(* IEC 61131-3 sources: Test-Git_ESME26/TestProgettoESME_26.fbsproj/PacDriveLib Migration/Motion/MultiCam/PDL_FB_MultiCam.fb.st^/PlcOpen, 3 files *)

(* ---- CallPLCopenFBs.meth.st ---- *)
METHOD PRIVATE CallPLCopenFBs : BOOL
VAR_INPUT
END_VAR

(*********************************************************************************************************************)
fbMoveAbsolute();

IF fbMoveAbsolute.Error THEN
	SetDiagOutput(	i_etDiag	:= GD.ET_Diag.UnexpectedProgramBehavior,
					i_etDiagExt := PDL_ET_DiagExt.UnexpectedFeedback,
					i_sMsg		:= CONCAT('MC_MoveAbsolute.ErrorID: ', PLCO.FC_EtResultToString(fbMoveAbsolute.ErrorID) ));
	fbMoveAbsolute.Execute := FALSE;

	q_xReady		:= FALSE;
	q_xSynActive	:= FALSE;
	q_xXLowEnd		:= FALSE;
	q_xXHighEnd		:= FALSE;
	q_xInWSWindow	:= FALSE;
	etState := ET_MulticamState.controllerStop;
END_IF

(*********************************************************************************************************************)
fbCamIn();

IF fbCamIn.Error THEN

	SetDiagOutput(	i_etDiag	:= GD.ET_Diag.UnexpectedProgramBehavior,
					i_etDiagExt := PDL_ET_DiagExt.UnexpectedFeedback,
					i_sMsg		:= CONCAT('MC_CamIn.ErrorID: ', PLCO.FC_EtResultToString(fbCamIn.ErrorID) ));

	fbCamIn.Execute := FALSE;
	q_xReady		:= FALSE;
	q_xSynActive	:= FALSE;
	q_xXLowEnd		:= FALSE;
	q_xXHighEnd		:= FALSE;
	q_xInWSWindow	:= FALSE;
	etState := ET_MulticamState.controllerStop;
END_IF

(*********************************************************************************************************************)
fbCamIn2();

IF fbCamIn2.Error THEN

	SetDiagOutput(	i_etDiag	:= GD.ET_Diag.UnexpectedProgramBehavior,
					i_etDiagExt := PDL_ET_DiagExt.UnexpectedFeedback,
					i_sMsg		:= CONCAT('MC_CamIn.ErrorID: ', PLCO.FC_EtResultToString(fbCamIn2.ErrorID) ));

	fbCamIn2.Execute := FALSE;
	q_xReady		:= FALSE;
	q_xSynActive	:= FALSE;
	q_xXLowEnd		:= FALSE;
	q_xXHighEnd		:= FALSE;
	q_xInWSWindow	:= FALSE;
	etState := ET_MulticamState.controllerStop;
END_IF

(*********************************************************************************************************************)

xCamInInSync :=    fbCamIn.InSync
			   AND NOT xCamIn2Active
			   OR  fbCamIn2.InSync
			   AND xCamIn2Active;

xCamInEndOfProfile :=      fbCamIn.EndOfProfile
					   AND NOT xCamIn2Active
					   OR  fbCamIn2.EndOfProfile
					   AND xCamIn2Active;

(* ---- SetPosition.meth.st ---- *)
METHOD PRIVATE SetPosition : BOOL
VAR_INPUT
	i_ifAxis		: MOIN.IF_Axis;
	i_lrPosition	: LREAL;
	i_xRelative		: BOOL;
END_VAR

VAR
	etSetPosResult				: PLCO.ET_Result;
END_VAR

SetPosition := TRUE;

fbSetPos( Execute		:= FALSE );
fbSetPos(	Axis		:= i_ifAxis,
			Execute		:= TRUE,
			Position	:= i_lrPosition,
			Relative	:= i_xRelative,
			ErrorId		=> etSetPosResult );

IF etSetPosResult <> PLCO.ET_Result.Ok THEN

	SetDiagOutput(	i_etDiag	:= GD.ET_Diag.UnexpectedProgramBehavior,
					i_etDiagExt := PDL_ET_DiagExt.UnexpectedFeedback,
					i_sMsg		:= CONCAT('MC_SetPosition: ', TO_STRING(etSetPosResult)));

	SetPosition := FALSE;//no success

	etState := ET_MulticamState.controllerStop;
END_IF

(* ---- StartCam.meth.st ---- *)
METHOD PRIVATE StartCam : BOOL
VAR_INPUT
	i_etBufferMode 			: PLCO.MC_Buffer_Mode;
	i_stMultiCamData		: PDL_ST_MultiCam;
	i_lrMasterStartPosition	: LREAL := 0;
	i_xPeriodic 			: BOOL := TRUE;
	i_etMasterStartMode		: PLCO.MC_Master_Start_Mode := PLCO.MC_Master_Start_Mode.Absolute;
	i_etSlaveStartMode		: PLCO.MC_Slave_Start_Mode := PLCO.MC_Slave_Start_Mode.RampIn;
	i_xInputVelocity		: BOOL := FALSE;
	i_etDirection			: PLCO.MC_Direction := PLCO.MC_Direction.ShortestWay;
END_VAR

IF xCamIn2Active THEN

	//camIn1
	//***********************************************************************************
	xCamIn2Active := FALSE;
	fbCamIn2( Execute := FALSE );

	IF i_xInputVelocity THEN
		fbCamIn.VelocityOffsetRampIn		:= i_lrWSVel;
		fbCamIn.AccelerationOffsetRampIn	:= i_lrWSAcc;
		fbCamIn.DecelerationOffsetRampIn	:= i_lrWSAcc;
		fbCamIn.JerkOffsetRampIn			:= i_lrWsJerk;
	ELSE
		IF ifDriveConfig <> 0 THEN
			IF ifDriveConfig.MaxVel <> 0 THEN
				fbCamIn.VelocityOffsetRampIn		:= ifDriveConfig.MaxVel;
			ELSE
				fbCamIn.VelocityOffsetRampIn		:= lrLimitMaxVel;
			END_IF

			IF ifDriveConfig.MaxAcc <> 0 THEN
				fbCamIn.AccelerationOffsetRampIn	:= ifDriveConfig.MaxAcc;
				fbCamIn.DecelerationOffsetRampIn	:= ifDriveConfig.MaxAcc;
			ELSE
				fbCamIn.AccelerationOffsetRampIn	:= lrLimitMaxAccDec;
				fbCamIn.DecelerationOffsetRampIn	:= lrLimitMaxAccDec;
			END_IF
		ELSE
			fbCamIn.VelocityOffsetRampIn		:= lrLimitMaxVel;
			fbCamIn.AccelerationOffsetRampIn	:= lrLimitMaxAccDec;
			fbCamIn.DecelerationOffsetRampIn	:= lrLimitMaxAccDec;
		END_IF
		fbCamIn.JerkOffsetRampIn			:= 0;
	END_IF

	fbCamIn(	Execute						:= TRUE,
				CamTableID					:= i_stMultiCamData,
				BufferMode					:= i_etBufferMode,
				Periodic					:= i_xPeriodic,
				MasterOffset				:= 0,
				SlaveOffset					:= 0,
				MasterScaling				:= 1,
				SlaveScaling				:= 1,
				MasterStartMode				:= i_etMasterStartMode,
				SlaveStartMode				:= i_etSlaveStartMode,
				RampInDirection				:= i_etDirection,
				MasterStartPosition			:= i_lrMasterStartPosition);

ELSE
	//camIn2
	//***********************************************************************************
	xCamIn2Active := TRUE;
	fbCamIn( Execute := FALSE );

	IF i_xInputVelocity THEN
		fbCamIn2.VelocityOffsetRampIn		:= i_lrWSVel;
		fbCamIn2.AccelerationOffsetRampIn	:= i_lrWSAcc;
		fbCamIn2.DecelerationOffsetRampIn	:= i_lrWSAcc;
		fbCamIn2.JerkOffsetRampIn			:= i_lrWsJerk;
	ELSE
		IF ifDriveConfig <> 0 THEN
			IF ifDriveConfig.MaxVel <> 0 THEN
				fbCamIn2.VelocityOffsetRampIn		:= ifDriveConfig.MaxVel;
			ELSE
				fbCamIn2.VelocityOffsetRampIn		:= lrLimitMaxVel;
			END_IF
			IF ifDriveConfig.MaxAcc <> 0 THEN
				fbCamIn2.AccelerationOffsetRampIn	:= ifDriveConfig.MaxAcc;
				fbCamIn2.DecelerationOffsetRampIn	:= ifDriveConfig.MaxAcc;
			ELSE
				fbCamIn2.AccelerationOffsetRampIn	:= lrLimitMaxAccDec;
				fbCamIn2.DecelerationOffsetRampIn	:= lrLimitMaxAccDec;
			END_IF
		ELSE
			fbCamIn.VelocityOffsetRampIn		:= lrLimitMaxVel;
			fbCamIn.AccelerationOffsetRampIn	:= lrLimitMaxAccDec;
			fbCamIn.DecelerationOffsetRampIn	:= lrLimitMaxAccDec;
		END_IF
		fbCamIn2.JerkOffsetRampIn			:= 0;
	END_IF

	fbCamIn2(	Execute						:= TRUE,
				CamTableID					:= i_stMultiCamData,
				BufferMode					:= i_etBufferMode,
				Periodic					:= i_xPeriodic,
				MasterOffset				:= 0,
				SlaveOffset					:= 0,
				MasterScaling				:= 1,
				SlaveScaling				:= 1,
				MasterStartMode				:= i_etMasterStartMode,
				SlaveStartMode				:= i_etSlaveStartMode,
				RampInDirection				:= i_etDirection,
				MasterStartPosition			:= i_lrMasterStartPosition);

END_IF
